Fanuc KAREL source: KT00510.KL

PROGRAM KT00510
%NOLOCKGROUP
VAR
  P1: XYZWPR
  P2: JOINTPOS
  OUT: XYZWPR
BEGIN
  P1.X = 1.0
  OUT = P1 : P2
END KT00510
